Fanuc KAREL source: KT00422.KL

PROGRAM KT00422
%NOLOCKGROUP
VAR
  P1: POSITION
  P2: JOINTPOS
  OUT: BOOLEAN
BEGIN
  OUT = P1 > P2
END KT00422
